(* IEC 61131-3 sources: trust-platform/crates/trust-runtime/tests/fixtures/oscat/core/src/16_logic_modules, 1 file *)

(* ---- tests.st ---- *)
TEST_PROGRAM oscat_logic_decoders_and_muxes_behave
VAR
    Dec2 : DEC_2;
    Dec4 : DEC_4;
    Dec8 : DEC_8;
    Selected2 : BOOL;
    Selected4 : BOOL;
END_VAR

Dec2(ENABLE := TRUE, A := FALSE);
ASSERT_TRUE(IN := Dec2.Q0);
ASSERT_FALSE(IN := Dec2.Q1);

Dec2(ENABLE := TRUE, A := TRUE);
ASSERT_FALSE(IN := Dec2.Q0);
ASSERT_TRUE(IN := Dec2.Q1);

Dec2(ENABLE := FALSE, A := TRUE);
ASSERT_FALSE(IN := Dec2.Q0);
ASSERT_FALSE(IN := Dec2.Q1);

Dec4(ENABLE := TRUE, A0 := TRUE, A1 := FALSE);
ASSERT_FALSE(IN := Dec4.Q0);
ASSERT_TRUE(IN := Dec4.Q1);
ASSERT_FALSE(IN := Dec4.Q2);
ASSERT_FALSE(IN := Dec4.Q3);

Dec4(ENABLE := TRUE, A0 := FALSE, A1 := TRUE);
ASSERT_FALSE(IN := Dec4.Q0);
ASSERT_FALSE(IN := Dec4.Q1);
ASSERT_TRUE(IN := Dec4.Q2);
ASSERT_FALSE(IN := Dec4.Q3);

Dec8(ENABLE := TRUE, A0 := TRUE, A1 := FALSE, A2 := TRUE);
ASSERT_FALSE(IN := Dec8.Q0);
ASSERT_FALSE(IN := Dec8.Q1);
ASSERT_FALSE(IN := Dec8.Q2);
ASSERT_FALSE(IN := Dec8.Q3);
ASSERT_FALSE(IN := Dec8.Q4);
ASSERT_TRUE(IN := Dec8.Q5);
ASSERT_FALSE(IN := Dec8.Q6);
ASSERT_FALSE(IN := Dec8.Q7);

Dec8(ENABLE := FALSE, A0 := TRUE, A1 := TRUE, A2 := TRUE);
ASSERT_FALSE(IN := Dec8.Q0);
ASSERT_FALSE(IN := Dec8.Q7);

Selected2 := MUX_2(D0 := FALSE, D1 := TRUE, A0 := FALSE);
ASSERT_FALSE(IN := Selected2);

Selected2 := MUX_2(D0 := FALSE, D1 := TRUE, A0 := TRUE);
ASSERT_TRUE(IN := Selected2);

Selected4 := MUX_4(D0 := FALSE, D1 := TRUE, D2 := TRUE, D3 := FALSE, A0 := FALSE, A1 := FALSE);
ASSERT_FALSE(IN := Selected4);

Selected4 := MUX_4(D0 := FALSE, D1 := TRUE, D2 := TRUE, D3 := FALSE, A0 := TRUE, A1 := FALSE);
ASSERT_TRUE(IN := Selected4);

Selected4 := MUX_4(D0 := FALSE, D1 := TRUE, D2 := TRUE, D3 := FALSE, A0 := FALSE, A1 := TRUE);
ASSERT_TRUE(IN := Selected4);

Selected4 := MUX_4(D0 := FALSE, D1 := TRUE, D2 := TRUE, D3 := FALSE, A0 := TRUE, A1 := TRUE);
ASSERT_FALSE(IN := Selected4);
END_TEST_PROGRAM

TEST_PROGRAM oscat_logic_bit_helpers_behave
VAR
    ByteBits : BYTE_TO_BITS;
    ByteValue : BYTE;
    DWordValue : DWORD;
    WordValue : WORD;
END_VAR

ASSERT_EQUAL(EXPECTED := INT#42, ACTUAL := BCDC_TO_INT(IN := BYTE#16#42));
ASSERT_EQUAL(EXPECTED := BYTE#16#42, ACTUAL := INT_TO_BCDC(IN := INT#42));

ASSERT_EQUAL(EXPECTED := INT#9, ACTUAL := BIT_COUNT(IN := DWORD#16#F0F00001));
ASSERT_TRUE(IN := BIT_OF_DWORD(IN := DWORD#16#10, N := INT#4));
ASSERT_FALSE(IN := BIT_OF_DWORD(IN := DWORD#16#10, N := INT#3));

ASSERT_EQUAL(EXPECTED := BYTE#8, ACTUAL := BIT_TOGGLE_B(IN := BYTE#0, POS := INT#3));
ASSERT_EQUAL(EXPECTED := WORD#16#1000, ACTUAL := BIT_TOGGLE_W(IN := WORD#0, POS := INT#12));
ASSERT_EQUAL(EXPECTED := DWORD#16#80000000, ACTUAL := BIT_TOGGLE_DW(IN := DWORD#0, POS := INT#31));

ByteValue := BYTE_OF_BIT(
    B0 := TRUE,
    B1 := FALSE,
    B2 := TRUE,
    B3 := FALSE,
    B4 := FALSE,
    B5 := TRUE,
    B6 := FALSE,
    B7 := TRUE
);
ASSERT_EQUAL(EXPECTED := BYTE#16#A5, ACTUAL := ByteValue);

ASSERT_EQUAL(EXPECTED := BYTE#16#AB, ACTUAL := BYTE_OF_DWORD(IN := DWORD#16#1234ABCD, N := BYTE#1));

ByteBits(IN := BYTE#16#A5);
ASSERT_TRUE(IN := ByteBits.B0);
ASSERT_FALSE(IN := ByteBits.B1);
ASSERT_TRUE(IN := ByteBits.B2);
ASSERT_TRUE(IN := ByteBits.B5);
ASSERT_TRUE(IN := ByteBits.B7);

ASSERT_EQUAL(EXPECTED := BYTE#8, ACTUAL := BYTE_TO_GRAY(IN := BYTE#15));
ASSERT_EQUAL(EXPECTED := BYTE#15, ACTUAL := GRAY_TO_BYTE(IN := BYTE#8));

ASSERT_TRUE(IN := CHECK_PARITY(IN := DWORD#1, P := TRUE));
ASSERT_FALSE(IN := CHECK_PARITY(IN := DWORD#1, P := FALSE));
ASSERT_FALSE(IN := PARITY(IN := DWORD#0));
ASSERT_TRUE(IN := PARITY(IN := DWORD#1));

DWordValue := DWORD_OF_BYTE(B3 := BYTE#16#12, B2 := BYTE#16#34, B1 := BYTE#16#AB, B0 := BYTE#16#CD);
ASSERT_EQUAL(EXPECTED := DWORD#16#1234ABCD, ACTUAL := DWordValue);

DWordValue := DWORD_OF_WORD(W1 := WORD#16#1234, W0 := WORD#16#ABCD);
ASSERT_EQUAL(EXPECTED := DWORD#16#1234ABCD, ACTUAL := DWordValue);

ASSERT_EQUAL(EXPECTED := DWORD#16#2345678F, ACTUAL := SHL1(IN := DWORD#16#12345678, N := INT#4));
ASSERT_EQUAL(EXPECTED := DWORD#16#F1234567, ACTUAL := SHR1(IN := DWORD#16#12345678, N := INT#4));

ASSERT_EQUAL(EXPECTED := WORD#16#3412, ACTUAL := SWAP_BYTE(IN := WORD#16#1234));
ASSERT_EQUAL(EXPECTED := DWORD#16#CDAB3412, ACTUAL := SWAP_BYTE2(IN := DWORD#16#1234ABCD));

WordValue := WORD_OF_BYTE(B1 := BYTE#16#12, B0 := BYTE#16#34);
ASSERT_EQUAL(EXPECTED := WORD#16#1234, ACTUAL := WordValue);

ASSERT_EQUAL(EXPECTED := WORD#16#ABCD, ACTUAL := WORD_OF_DWORD(IN := DWORD#16#1234ABCD, N := BYTE#0));
ASSERT_EQUAL(EXPECTED := WORD#16#1234, ACTUAL := WORD_OF_DWORD(IN := DWORD#16#1234ABCD, N := BYTE#1));
END_TEST_PROGRAM

TEST_PROGRAM oscat_logic_bit_load_helpers_behave
ASSERT_EQUAL(EXPECTED := BYTE#8, ACTUAL := BIT_LOAD_B(IN := BYTE#0, VAL := TRUE, POS := INT#3));
ASSERT_EQUAL(EXPECTED := BYTE#0, ACTUAL := BIT_LOAD_B(IN := BYTE#8, VAL := FALSE, POS := INT#3));
ASSERT_EQUAL(EXPECTED := BYTE#14, ACTUAL := BIT_LOAD_B2(I := BYTE#0, VALUE := TRUE, P := INT#1, N := INT#3));
ASSERT_EQUAL(EXPECTED := BYTE#16#E3, ACTUAL := BIT_LOAD_B2(I := BYTE#16#FF, VALUE := FALSE, P := INT#2, N := INT#3));

ASSERT_EQUAL(EXPECTED := WORD#16#1000, ACTUAL := BIT_LOAD_W(IN := WORD#0, VAL := TRUE, POS := INT#12));
ASSERT_EQUAL(EXPECTED := WORD#0, ACTUAL := BIT_LOAD_W(IN := WORD#16#1000, VAL := FALSE, POS := INT#12));
ASSERT_EQUAL(EXPECTED := WORD#16#01F0, ACTUAL := BIT_LOAD_W2(I := WORD#0, VALUE := TRUE, P := INT#4, N := INT#5));
ASSERT_EQUAL(EXPECTED := WORD#16#FE0F, ACTUAL := BIT_LOAD_W2(I := WORD#16#FFFF, VALUE := FALSE, P := INT#4, N := INT#5));

ASSERT_EQUAL(EXPECTED := DWORD#16#80000000, ACTUAL := BIT_LOAD_DW(IN := DWORD#0, VAL := TRUE, POS := INT#31));
ASSERT_EQUAL(EXPECTED := DWORD#0, ACTUAL := BIT_LOAD_DW(IN := DWORD#16#80000000, VAL := FALSE, POS := INT#31));
ASSERT_EQUAL(EXPECTED := DWORD#16#0000FF00, ACTUAL := BIT_LOAD_DW2(I := DWORD#0, VALUE := TRUE, P := INT#8, N := INT#8));
ASSERT_EQUAL(EXPECTED := DWORD#16#FFFF00FF, ACTUAL := BIT_LOAD_DW2(I := DWORD#16#FFFFFFFF, VALUE := FALSE, P := INT#8, N := INT#8));
END_TEST_PROGRAM

TEST_PROGRAM oscat_logic_bit_cast_and_reflection_helpers_behave
VAR
    PositiveInfinity : REAL;
    NegativeInfinity : REAL;
    NotANumber : REAL;
END_VAR

ASSERT_EQUAL(EXPECTED := DWORD#16#3FC00000, ACTUAL := REAL_TO_DW(X := REAL#1.5));
ASSERT_NEAR(EXPECTED := REAL#1.5, ACTUAL := DW_TO_REAL(X := DWORD#16#3FC00000), DELTA := REAL#0.0001);

ASSERT_EQUAL(EXPECTED := DWORD#16#19, ACTUAL := REFLECT(VALUE := DWORD#16#13, L := INT#5));
ASSERT_EQUAL(EXPECTED := BYTE#16#69, ACTUAL := REVERSE(IN := BYTE#16#96));

ASSERT_EQUAL(EXPECTED := BYTE#16#00, ACTUAL := CHK_REAL(X := REAL#0.0));

PositiveInfinity := DWORD_TO_REAL(DWORD#16#7F800000);
NegativeInfinity := DWORD_TO_REAL(DWORD#16#FF800000);
NotANumber := DWORD_TO_REAL(DWORD#16#7FC00000);

ASSERT_EQUAL(EXPECTED := BYTE#16#20, ACTUAL := CHK_REAL(X := PositiveInfinity));
ASSERT_EQUAL(EXPECTED := BYTE#16#40, ACTUAL := CHK_REAL(X := NegativeInfinity));
ASSERT_EQUAL(EXPECTED := BYTE#16#80, ACTUAL := CHK_REAL(X := NotANumber));
END_TEST_PROGRAM

TEST_PROGRAM oscat_logic_crc_gen_behaves
VAR
    Data : ARRAY[0..3] OF BYTE;
    Checksum : DWORD;
END_VAR

Data[0] := BYTE#1;
Data[1] := BYTE#2;
Data[2] := BYTE#3;
Data[3] := BYTE#4;

Checksum := CRC_GEN(
    PT := ADR(Data),
    SIZE := INT#4,
    PL := INT#8,
    PN := DWORD#16#07,
    INIT := DWORD#0,
    REV_IN := FALSE,
    REV_OUT := FALSE,
    XOR_OUT := DWORD#0
);
ASSERT_EQUAL(EXPECTED := DWORD#16#E3, ACTUAL := Checksum);
END_TEST_PROGRAM

TEST_PROGRAM oscat_logic_matrix_helpers_behave
VAR
    PressOnly : MATRIX;
    WithRelease : MATRIX;
END_VAR

PressOnly(X1 := TRUE, X2 := FALSE, X3 := FALSE, X4 := FALSE, X5 := FALSE, Release := FALSE);
ASSERT_TRUE(IN := PressOnly.TP);
ASSERT_EQUAL(EXPECTED := BYTE#16#81, ACTUAL := PressOnly.CODE);

PressOnly(X1 := FALSE, X2 := FALSE, X3 := FALSE, X4 := FALSE, X5 := FALSE, Release := FALSE);
ASSERT_FALSE(IN := PressOnly.TP);
PressOnly(X1 := FALSE, X2 := FALSE, X3 := FALSE, X4 := FALSE, X5 := FALSE, Release := FALSE);
ASSERT_FALSE(IN := PressOnly.TP);
PressOnly(X1 := FALSE, X2 := FALSE, X3 := FALSE, X4 := FALSE, X5 := FALSE, Release := FALSE);
ASSERT_FALSE(IN := PressOnly.TP);
PressOnly(X1 := FALSE, X2 := FALSE, X3 := FALSE, X4 := FALSE, X5 := FALSE, Release := FALSE);
ASSERT_FALSE(IN := PressOnly.TP);
ASSERT_EQUAL(EXPECTED := BYTE#0, ACTUAL := PressOnly.CODE);

WithRelease(X1 := FALSE, X2 := TRUE, X3 := FALSE, X4 := FALSE, X5 := FALSE, Release := TRUE);
ASSERT_TRUE(IN := WithRelease.TP);
ASSERT_EQUAL(EXPECTED := BYTE#16#82, ACTUAL := WithRelease.CODE);

WithRelease(X1 := FALSE, X2 := FALSE, X3 := FALSE, X4 := FALSE, X5 := FALSE, Release := TRUE);
ASSERT_FALSE(IN := WithRelease.TP);
WithRelease(X1 := FALSE, X2 := FALSE, X3 := FALSE, X4 := FALSE, X5 := FALSE, Release := TRUE);
ASSERT_FALSE(IN := WithRelease.TP);
WithRelease(X1 := FALSE, X2 := FALSE, X3 := FALSE, X4 := FALSE, X5 := FALSE, Release := TRUE);
ASSERT_FALSE(IN := WithRelease.TP);
WithRelease(X1 := FALSE, X2 := FALSE, X3 := FALSE, X4 := FALSE, X5 := FALSE, Release := TRUE);
ASSERT_TRUE(IN := WithRelease.TP);
ASSERT_EQUAL(EXPECTED := BYTE#16#02, ACTUAL := WithRelease.CODE);
END_TEST_PROGRAM

TEST_PROGRAM oscat_logic_pin_code_helpers_behave
VAR
    Door : PIN_CODE;
END_VAR

Door(CB := BYTE#49, E := TRUE, PIN := '12');
ASSERT_FALSE(IN := Door.TP);
Door(CB := BYTE#50, E := TRUE, PIN := '12');
ASSERT_TRUE(IN := Door.TP);

Door(CB := BYTE#50, E := TRUE, PIN := '12');
ASSERT_FALSE(IN := Door.TP);
Door(CB := BYTE#49, E := TRUE, PIN := '12');
ASSERT_FALSE(IN := Door.TP);
Door(CB := BYTE#50, E := TRUE, PIN := '12');
ASSERT_TRUE(IN := Door.TP);
END_TEST_PROGRAM
